FUNCTION_BLOCK FB_Example
VAR PERSISTENT
	persist_int 	: INT;
	persist_str 	: T_MaxString;
	persist_float	: REAL;
END_VAR
VAR RETAIN
	retain_int 		: INT;
	retain_str 		: T_MaxString;
	retain_float	: REAL;
END_VAR
VAR 
	non_per		: INT;
	non_per2	: LREAL;
	timer		: TON;
END_VAR

END_FUNCTION_BLOCK

(* stored: Version 1.1.0.1
   POU FB_Example: Id {835cf410-ead8-48b0-85bf-3947854c84b8}, SpecialFunc None *)
